(*
This paragraph is not part of the list.

- This is the first bullet list item.  The blank line above the
  first list item is required; blank lines between list items
  (such as below this paragraph) are optional.

  - This is a sublist. The bullet lines up with the left edge
    of the text blocks above. A sublist is a new list so
    requires a blank line above. A blank line below is optional.

  - This is a sublist. The bullet lines up with the left edge
    of the text blocks above. A sublist is a new list so
    requires a blank line above. A blank line below is optional.

- This is the second item of the main list.

- This is the third item of the main list.

This paragraph is not part of the list.
*)

FUNCTION_BLOCK FB_Libdoc_UnorderedEnumerationList
VAR_INPUT
    nVarA : INT;
    nVarB : INT;
END_VAR
VAR_OUTPUT
    nSum : INT;
END_VAR
VAR
END_VAR

END_FUNCTION_BLOCK

(* stored: Version 1.1.0.1, ProductVersion 3.1.4022.17
   POU FB_Libdoc_UnorderedEnumerationList: Id {c5ffe2a0-6a14-48ae-9899-29dd8c6aec50}, SpecialFunc None *)
